(* ================================================================= *)
(*  类型名称：ST_SingleLayer                                          *)
(*  功能描述：单层输送机数据结构体 (FB_1002 通过 VAR_IN_OUT 整块传递)  *)
(*  版本号：V1.0.0 (2026-10-24, DJ-2026-005 新设计)                    *)
(*                                                                     *)
(*  依据：接口文档_INT.md 4.5；层号 1 = 最下层                         *)
(*  遵循规范：LSP-905 SCL编程规范                                      *)
(* ================================================================= *)

TYPE ST_SingleLayer
STRUCT
    (* ------------------ 传感器输入 ------------------ *)
    bPreBlock               : BOOL;     // 阻挡前到位传感器
    bPick1                  : BOOL;     // 边框取料位接近开关 1
    bPick2                  : BOOL;     // 边框取料位接近开关 2
    bFull1                  : BOOL;     // 边框满料检测 1
    bFull2                  : BOOL;     // 边框满料检测 2
    bBlkUp1                 : BOOL;     // 阻挡气缸上位 1
    bBlkUp2                 : BOOL;     // 阻挡气缸上位 2
    bBlkDn1                 : BOOL;     // 阻挡气缸下位 1
    bBlkDn2                 : BOOL;     // 阻挡气缸下位 2
    bSepUp1                 : BOOL;     // 分料气缸上位 1
    bSepUp2                 : BOOL;     // 分料气缸上位 2
    bSepDn1                 : BOOL;     // 分料气缸下位 1
    bSepDn2                 : BOOL;     // 分料气缸下位 2

    (* ------------------ 命令输入 ------------------ *)
    bInitReq                : BOOL;     // 初始化请求 (回原点预处理期间)
    bAutoRun                : BOOL;     // 自动运行
    bHold                   : BOOL;     // 本层保持 (暂停 / 本层报警 / 全局 Hold)
    bReset                  : BOOL;     // 异常停机 (M8 或进手动)
    bSafeZone               : BOOL;     // 取料机构在安全区
    bPickDone               : BOOL;     // 本层取料完成 (来自取放料, 本层对本层)
    bStopPending            : BOOL;     // 停止请求 (本循环结束后不再开新循环)

    (* ------------------ 命令输出 ------------------ *)
    bBlockDown              : BOOL;     // 阻挡下降命令 (ON = 下降放行, OFF = 升起)
    bSepDown                : BOOL;     // 分料下降命令 (ON = 下降压料, OFF = 升起)
    bFwd                    : BOOL;     // 输送正转
    bRev                    : BOOL;     // 输送反转
    bSlow                   : BOOL;     // 输送慢速 (只在正转或反转有效时才输出)

    (* ------------------ 状态输出 ------------------ *)
    bReady                  : BOOL;     // 准备完成
    bRequest                : BOOL;     // 请求取料
    bAtRest                 : BOOL;     // 静止点 (步 0), 供停止收尾判断
    iStep                   : INT;      // 当前步 (供 HMI / 测试)

    (* ------------------ 双向 ------------------ *)
    bUnload                 : BOOL;     // 退料 (HMI 置位, 4 层准备完成后由 FB_1007 清除)

    (* ------------------ 报警触发 ------------------ *)
    // [0..7] 阻挡上 1/上 2/下 1/下 2, 分料上 1/上 2/下 1/下 2 (对应 F34~F41 + 8 x (层号-1))
    // [8]    缺料 (对应 F103 - (层号-1))
    arrTrig                 : ARRAY[1..9] OF BOOL;      // 报警触发: [1..8] 气缸位置 (F34 起, 每层 +8), [9] 缺料 (F103 起, 每高一层 -1)
END_STRUCT
END_TYPE
